FUNCTION_BLOCK T_SafeOr_Tests EXTENDS TcUnit.FB_TestSuite
VAR
    // Test_AnyConnectedInputTrueGivesRun
    group_1 : T_SafeGroup;
    fb_1 : T_SafeOr(group := group_1);
    // Test_AllFalseGivesSafe
    group_2 : T_SafeGroup;
    fb_2 : T_SafeOr(group := group_2);
    // Test_OneConnectedInputIsRefused
    group_3 : T_SafeGroup;
    fb_3 : T_SafeOr(group := group_3);
END_VAR

Test_AnyConnectedInputTrueGivesRun();
Test_AllFalseGivesSafe();
Test_OneConnectedInputIsRefused();

METHOD PRIVATE Test_AllFalseGivesSafe
TcUnit.TEST(__POUNAME());
// act
group_2(Run := TRUE);
fb_2(OrIn1 := FALSE, OrIn2 := FALSE);
// assert
AssertEquals_BOOL(Expected := FALSE, Actual := fb_2.OrOut, Message := 'output off when all connected inputs are 0');
AssertEquals_BYTE(Expected := TO_BYTE(E_SafeFbState.Safe), Actual := fb_2.State, Message := 'state SAFE');
TEST_FINISHED_NAMED(__POUNAME());
END_METHOD

METHOD PRIVATE Test_AnyConnectedInputTrueGivesRun
TcUnit.TEST(__POUNAME());
// act
group_1(Run := TRUE);
fb_1(OrIn1 := FALSE, OrIn2 := TRUE);
// assert
AssertEquals_BOOL(Expected := TRUE, Actual := fb_1.OrOut, Message := 'output on when any connected input is 1');
TEST_FINISHED_NAMED(__POUNAME());
END_METHOD

METHOD PRIVATE Test_OneConnectedInputIsRefused
TcUnit.TEST(__POUNAME());
// arrange / act: OrIn1 is the only connected input, which the Safety Editor refuses
group_3(Run := TRUE);
fb_3(OrIn1 := TRUE);
group_3(Run := TRUE);
fb_3(OrIn1 := TRUE);
// assert
AssertEquals_BOOL(Expected := TRUE, Actual := fb_3.Error, Message := 'configuration error reported');
AssertEquals_BYTE(Expected := TO_BYTE(E_SafeFbState.Error), Actual := fb_3.State, Message := 'state ERROR');
AssertEquals_WORD(Expected := WORD#16#8000, Actual := fb_3.Diag, Message := 'diag bit 15 configuration refused');
AssertEquals_BOOL(Expected := FALSE, Actual := fb_3.OrOut, Message := 'OrOut stays at its safe value');
AssertEquals_BOOL(Expected := TRUE, Actual := group_3.FbErr, Message := 'the group sees an FB error');
// act: ErrAck 0 -> 1 -> 0 does not clear a configuration error
group_3(Run := TRUE, ErrAck := TRUE);
fb_3(OrIn1 := TRUE);
group_3(Run := TRUE, ErrAck := TRUE);
fb_3(OrIn1 := TRUE);
group_3(Run := TRUE, ErrAck := FALSE);
fb_3(OrIn1 := TRUE);
AssertEquals_BOOL(Expected := TRUE, Actual := fb_3.Error, Message := 'error not acknowledged');
AssertEquals_WORD(Expected := WORD#16#8000, Actual := fb_3.Diag, Message := 'diag bit 15 kept');
TEST_FINISHED_NAMED(__POUNAME());
END_METHOD

END_FUNCTION_BLOCK

(* stored: Version 1.1.0.1
   POU T_SafeOr_Tests: Id {04c9cafe-7788-59b6-a714-e1b30ac42516}, SpecialFunc None
   Method Test_AllFalseGivesSafe: Id {7edfe92d-179f-53fa-be6a-5be0f61c49b9}
   Method Test_AnyConnectedInputTrueGivesRun: Id {cf343ecd-ee19-52cd-bcab-51e8b478f6eb}
   Method Test_OneConnectedInputIsRefused: Id {a50db1bc-ec9d-4e63-bba1-7dce482328e2} *)
